Fanuc KAREL source: kx00031.KL

-- PROVISIONAL review KL for V1013-1; original PC SHA256 9b8e3ec29dd3350a8c49971cdc9fc36ab5f1c4dacceee4b564bcf002400eba6a
-- Incomplete behavior may be omitted. Consult companion uncertainty JSON. Do not deploy.
PROGRAM KX00031
%NOLOCKGROUP
VAR
  I : INTEGER
  J : INTEGER
  B : BOOLEAN
  F : FILE
  S : STRING[80]
-- UNRESOLVED_DECL P type=000102
BEGIN
  -- UNRESOLVED_PC offsets 5-12; opcodes 9D,23
  -- UNRESOLVED_PC offsets 17-21; opcodes 7F
END KX00031
